Fanuc KAREL source: KT00195.KL

PROGRAM KT00195
%NOLOCKGROUP
VAR
  B1: BOOLEAN
  I2: INTEGER
  OUT: BOOLEAN
BEGIN
  B1 = TRUE
    I2 = 3
  OUT = B1 AND I2
END KT00195
